Staubli VAL3: setframemode.pgx

public program setframemode()
  local num l_i
begin
  $jogMode(2)
  for l_i = 0 to size(sShowType)-1
    sShowType[l_i]=sCartisiam[l_i]
  endFor
end
